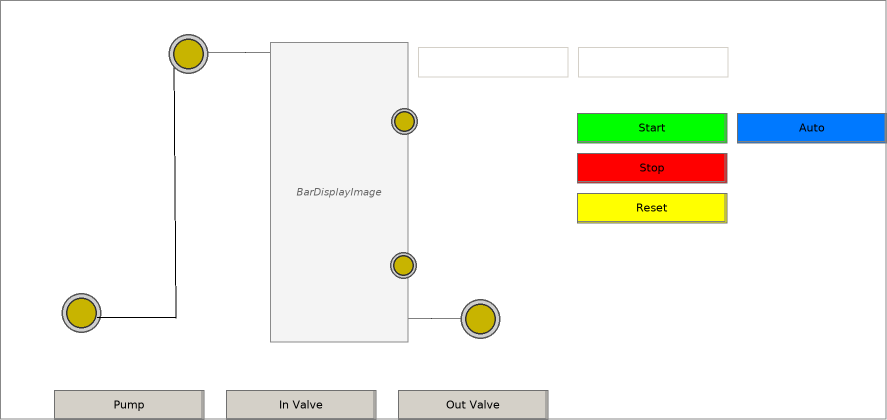
VISUALIZATION TankVisual  // 887x420
    Line (474,319) (389,318)
    Line (288,53) (203,52)
    Rectangle (270,42 138x300)
    BarDisplayImage (270,42 138x300), value: GVL_HMI.Tank1.rLevel, style: BarDisplayImage-Gray, scale format: %.1f, scale 0..100
    Lamp1 (453,296 55x46), variable: GVL_HMI.Tank1.bPB_ValveOut, style: Lamp-Lamp1-Yellow
    Lamp1 (54,290 55x46), variable: GVL_HMI.Tank1.bPB_Pump, style: Lamp-Lamp1-Yellow
    Lamp1 (389,106 31x31), variable: MAIN.bSensHIGH, style: Lamp-Lamp1-Yellow
    Lamp1 (388,250 31x31), variable: MAIN.bSensLOW, style: Lamp-Lamp1-Yellow
    Button (577,113 150x30), "Start", pressed state: GVL_HMI.Tank1.bStart
    Button (737,113 150x30), "Auto", pressed state: GVL_HMI.Tank1.bAutoMode
        toggle GVL_HMI.Tank1.bAutoMode p2164770859=TRUE
    Button (54,390 150x30), "Pump", input disabled if: GVL_HMI.Tank1.bAutoMode
        tap GVL_HMI.Tank1.bPB_Pump
        toggle GVL_HMI.Tank1.bPB_Pump
    Button (226,390 150x30), "In Valve", input disabled if: GVL_HMI.Tank1.bAutoMode
        toggle GVL_HMI.Tank1.bPB_ValveIn
    Button (398,390 150x30), "Out Valve", input disabled if: GVL_HMI.Tank1.bAutoMode
        toggle GVL_HMI.Tank1.bPB_ValveOut
    Line (97,317) (176,317)
    Line (176,318) (174,58)
    Lamp1 (161,31 55x46), variable: GVL_HMI.Tank1.bPB_ValveIn, style: Lamp-Lamp1-Yellow
    Button (577,193 150x30), "Reset", pressed state: GVL_HMI.Tank1.bReset
    Button (577,153 150x30), "Stop", pressed state: GVL_HMI.Tank1.bStop
    Textfield (418,47 150x30), text variable: GVL_HMI.Tank1.eState
    Textfield (578,47 150x30), text variable: GVL_HMI.Tank1.eState
END_VISUALIZATION

(* stored: Version 1.1.0.1
   Visu TankVisual: Id {c6d20605-bb37-41cb-b812-dff7e04dacfa} *)
